FUNCTION_BLOCK FB_Homing_Modulo EXTENDS FB_Homing_Base IMPLEMENTS I_MotionSequence
VAR_INPUT
    ReferencePosition : LREAL := 0.0;
END_VAR
VAR
    fbMcHome          : MC_Home;
    fbMoveAbs         : MC_MoveAbsolute;
    fbSetPosition     : MC_SetPosition; 
    _HomingVelocity   : LREAL := 50.0;
    _TargetPos        : LREAL := 0.0;
END_VAR

METHOD Abort
VAR_INPUT
END_VAR
IF _Axis <> 0 THEN
    fbMcHome(Axis := _Axis.Axis, Execute := FALSE);
    fbMoveAbs(Axis := _Axis.Axis, Execute := FALSE);
    fbSetPosition(Axis := _Axis.Axis, Execute := FALSE); 
END_IF

SUPER^.Abort();
END_METHOD

METHOD CyclicLogic
VAR
    lrCurrentPos : LREAL;
    lrRemainder  : LREAL;
END_VAR


CASE nStep OF
    0: 
        fbMcHome(Axis := _Axis.Axis, Execute := FALSE);
        fbMoveAbs(Axis := _Axis.Axis, Execute := FALSE);
        fbSetPosition(Axis := _Axis.Axis, Execute := FALSE); 

		10: 
			IF _Axis.Axis.Status.Homed THEN
				ADSLOGSTR(ADSLOG_MSGTYPE_ERROR, '6. HomingModulo [Step 10] -> AxisQ juz Homed=TRUE, ide do 15', '');
				nStep := 15;
			ELSE
				IF NOT fbMcHome.Busy THEN
					ADSLOGSTR(ADSLOG_MSGTYPE_ERROR, '6. HomingModulo [Step 10] -> start MC_Home(MC_Direct)', '');
				END_IF
				fbMcHome(
					Axis        := _Axis.Axis, 
					Execute     := TRUE, 
					Position    := ReferencePosition,
					HomingMode  := MC_Direct
				);
				
				IF fbMcHome.Done THEN
					ADSLOGSTR(ADSLOG_MSGTYPE_ERROR, '6a. HomingModulo [Step 10] -> MC_Home DONE', '');
					fbMcHome(Axis := _Axis.Axis, Execute := FALSE);
					nStep := 15;
				ELSIF fbMcHome.Error THEN
					ADSLOGSTR(ADSLOG_MSGTYPE_ERROR, 'BLAD HomingModulo [Step 10] -> MC_Home ErrorID: %s', UDINT_TO_STRING(fbMcHome.ErrorID));
					_bBusy    := FALSE;
					_bError   := TRUE;
					_bErrorID := fbMcHome.ErrorID;
					nStep     := 0;
				END_IF
			END_IF
		
15:
        lrCurrentPos := _Axis.Axis.NcToPlc.ActPos;
        lrRemainder  := lrCurrentPos - DINT_TO_LREAL(LREAL_TO_DINT(lrCurrentPos / 360.0)) * 360.0;
        _TargetPos   := lrRemainder; // Zapis do zmiennej instancyjnej FB (nie ginie w kolejnym cyklu!)
        ADSLOGSTR(ADSLOG_MSGTYPE_ERROR, '7. HomingModulo [Step 15] -> ActPos=%s', LREAL_TO_STRING(lrCurrentPos));
        ADSLOGSTR(ADSLOG_MSGTYPE_ERROR, '7a. HomingModulo [Step 15] -> zapisano _TargetPos=%s', LREAL_TO_STRING(_TargetPos));
        nStep        := 20;

    20:
        IF NOT fbSetPosition.Busy THEN
            ADSLOGSTR(ADSLOG_MSGTYPE_ERROR, '8. HomingModulo [Step 20] -> start MC_SetPosition na: %s', LREAL_TO_STRING(_TargetPos));
        END_IF

        fbSetPosition(
            Axis     := _Axis.Axis,
            Execute  := TRUE,
            Position := _TargetPos, // Tu jest +90.0°, więc NC wie, że nóż jest 90° od oryginalnego 0°
            Mode     := FALSE
        );
        
        IF fbSetPosition.Done THEN
            ADSLOGSTR(ADSLOG_MSGTYPE_ERROR, '9. HomingModulo [Step 20] -> MC_SetPosition DONE', '');
            fbSetPosition(Axis := _Axis.Axis, Execute := FALSE);
            nStep := 30;
        ELSIF fbSetPosition.Error THEN
            ADSLOGSTR(ADSLOG_MSGTYPE_ERROR, 'BLAD HomingModulo [Step 20] -> MC_SetPosition ErrorID: %s', UDINT_TO_STRING(fbSetPosition.ErrorID));
            _bBusy    := FALSE;
            _bError   := TRUE;
            _bErrorID := fbSetPosition.ErrorID;
            nStep     := 0;
        END_IF

    30: 
        IF NOT fbMoveAbs.Busy THEN
            ADSLOGSTR(ADSLOG_MSGTYPE_ERROR, '10. HomingModulo [Step 30] -> start MC_MoveAbsolute do 0.0', '');
        END_IF

        fbMoveAbs(
            Axis      := _Axis.Axis,
            Execute   := TRUE,
            Position  := 0.0, // Fizyczny obrót z +90.0° na oryginalne 0.0° (ruch o -90°)
            Velocity  := _HomingVelocity
        );
        
        IF fbMoveAbs.Done THEN
            ADSLOGSTR(ADSLOG_MSGTYPE_ERROR, '11. HomingModulo [Step 30] -> MC_MoveAbsolute DONE (os na 0.0)', '');
            fbMoveAbs(Axis := _Axis.Axis, Execute := FALSE);
            nStep := 40; 
        ELSIF fbMoveAbs.Error THEN
            ADSLOGSTR(ADSLOG_MSGTYPE_ERROR, 'BLAD HomingModulo [Step 30] -> MC_MoveAbsolute ErrorID: %s', UDINT_TO_STRING(fbMoveAbs.ErrorID));
            _bBusy    := FALSE;
            _bError   := TRUE;
            _bErrorID := fbMoveAbs.ErrorID;
            nStep     := 0;
        END_IF
        
    40: 
        _bBusy := FALSE;
        _bDone := TRUE; 
        nStep  := 0;
END_CASE
END_METHOD

PROPERTY HomingVelocity : LREAL
GET
HomingVelocity := _HomingVelocity;
END_GET
SET
_HomingVelocity := HomingVelocity;
END_SET
END_PROPERTY

END_FUNCTION_BLOCK

(* stored: Version 1.1.0.1, ProductVersion 3.1.4024.15
   POU FB_Homing_Modulo: Id {398b7abf-73ed-4a8a-a3c8-2f04463db183}, SpecialFunc None
   Method Abort: Id {3c597dbe-7762-4228-aa6b-316da941959e}
   Method CyclicLogic: Id {afe30813-6e1e-4130-8cfc-c80e37369084}
   Property HomingVelocity: Id {551cdd69-c6cb-47ff-b9b7-6792dba04d4f}
   Get Get: Id {8b56f16c-648b-4463-a280-406b1f5b5952}
   Set Set: Id {324ec116-8e07-4c79-9459-8dcef86359a2} *)
